Staubli VAL3: _clickAlarmAck.pgx

program _clickAlarmAck()
begin
  rs:_sRobotStatus="收到页面点击清除报错!"
  rs:bAlarmAck=true
  delay(0.1)
  rs:bAlarmAck=false
end
